Fanuc KAREL source: kt00524.KL

-- PROVISIONAL review KL for V940-1; original PC SHA256 aaa6ae2c1c3a5b7d4d7b1ff1a45d531f53125e5289bfede18ba29a6fa5f6a12b
-- Incomplete behavior may be omitted. Consult companion uncertainty JSON. Do not deploy.
PROGRAM KT00524
%NOLOCKGROUP
-- UNRESOLVED_DECL P1 type=000106
-- UNRESOLVED_DECL P2 type=000106
-- UNRESOLVED_DECL OUT type=000101
BEGIN
  -- V9_ZERO_TABLE_METADATA_HINT layout=0001; no indexed target words; source/name/runtime held
  -- UNRESOLVED_PC offsets 5-20; opcodes 2E,22,32,35
  -- UNRESOLVED_PC offsets 25-40; opcodes 2E,22,32,35
  -- UNRESOLVED_PC offsets 45-60; opcodes 2E,22,32,35
  -- UNRESOLVED_PC offsets 65-80; opcodes 2E,22,32,35
  -- UNRESOLVED_PC offsets 85-119; opcodes 49,7E,49,7E,60,4A
  -- UNRESOLVED_PC offsets 124-128; opcodes 7F
END KT00524
